{attribute 'OPC.UA.DA.StructuredType' := '1'}
TYPE ST_HeatPumpAirState :
STRUCT
	bError	: BOOL;
	bCommunicationError : BOOL;
	bPlantMode : UDINT;
	bSystemMode : UDINT;
	fAmbientTemperature : REAL;
	fFeedTemperature : REAL;
	fReturnTemperature : REAL;
	fBufferTemperatureTop : REAL;
	fBufferTemperatureBottom : REAL;
	fPowersetpoint : REAL;
	fOperatingHours	 : UDINT;
	nCycles : UDINT;
	
END_STRUCT
END_TYPE

(* stored: Version 1.1.0.1
   DUT ST_HeatPumpAirState: Id {3a548344-f1e9-4850-bf9e-c5c25b0c4b0f} *)
